(* IEC 61131-3 sources: daoli-st-library/DL_Process (part 24) *)

(* ---- FB_DL_CartonErectSeq.st ---- *)
(*==============================================================================
 * 组件名称 (Component)  : FB_DL_CartonErectSeq
 * 所属子库 (Sublibrary) : DL_Process
 * 当前版本 (Version)    : 1.0.0
 * 兼容性 (Platform)     : CODESYS 3.5 / TwinCAT 3 / 汇川 InoProShop / Machine Expert
 *                         仅依赖纯 IEC 61131-3 标准元素，零厂商方言
 * 功能描述 (Function)   : 开箱机顺控四相：吸箱 → 成型 → 折底 → 输送，含卡箱检测，
 *                         单相超时（tStepMax 默认 5 s）监视；反馈缺失一律进 ERR
 *                         并锁存卡箱（不跳相）；PICK 相真空超时先释放真空再报错；
 *                         CASE 含 ELSE 安全态（全输出 FALSE）；复位退 IDLE。
 * 溯源 (Origin)         : 道莅 clean-room 防御性实现
 * 本文件内含 (Contains) : TYPE E_DL_ErectPhase / TYPE E_DL_ErectErr /
 *                         FUNCTION_BLOCK FB_DL_CartonErectSeq
 * 依赖 (Depends)        : 无 DL_ 内部依赖；Standard.library TON/R_TRIG 实例
 * 红线自检 (Redline)    : 无外部全局变量、无硬件地址直引 ｜ 全变量中英双语同行注释
 *                         相超时用状态判定（TON.Q + 相枚举），非单拍标志 ｜
 *                         枚举成员全部显式赋值 ｜ TON/R_TRIG 每周期无条件调用 ｜
 *                         CASE 含 ELSE 兜底至安全态 ｜ 无占位词 ｜ 超时引脚带单位
 * 错误码表 (Codes)      : 16#0005_041C IDLE（或 DONE 等待下一循环，共用反证句）
 *                         16#0005_041D PICK（吸箱相）
 *                         16#0005_041E FORM（成型相）
 *                         16#0005_041F FLAP（折底相，EJECT 输送段共用反证句）
 *                         16#0005_0420 ERR（含相超时定位，定位另由 eJamPhase 输出）
 * 修订历史 (Revision)   : 2026-11-17  v1.0.0  首版入库 · R27 · 阶段三批 4
 * 验收向量 (Acceptance) : bStart → PICK（真空指令置位）→ bVacuumOk → FORM → bBoxFormed
 *                         → FLAP → bFlapClosed → EJECT → DONE；PICK 相 tStepMax 内
 *                         无 bVacuumOk → ERR + bJam + 真空撤 + eJamPhase=PICK
 *============================================================================*)

(*-----------------------------------------------------------------------------
 * 枚举: E_DL_ErectPhase（归属 DL_Process，开箱顺控相）
 *----------------------------------------------------------------------------*)
TYPE E_DL_ErectPhase :
(
    ePhaseIdle  := 0,    // 空闲待启动 / Idle, waiting for a start
    ePhasePick  := 10,   // 吸箱相（真空建立）/ Pick phase, vacuum build-up
    ePhaseForm  := 20,   // 成型相 / Forming phase
    ePhaseFlap  := 30,   // 折底相 / Flap-closing phase
    ePhaseEject := 40,   // 输送相（定时完成）/ Eject phase, timed
    ePhaseDone  := 50,   // 循环完成（等待下一循环）/ Cycle done, waiting for the next
    ePhaseErr   := 99    // 故障相（卡箱锁存）/ Error phase, jam latched
);
END_TYPE

(*-----------------------------------------------------------------------------
 * 枚举: E_DL_ErectErr（归属 DL_Process，与 FB_DL_CartonErectSeq 同文件）
 *----------------------------------------------------------------------------*)
TYPE E_DL_ErectErr :
(
    eIdle   := 16#0005_041C,   // IDLE（含 DONE 等待态）/ Idle or done-waiting
    ePick   := 16#0005_041D,   // PICK 相（吸箱）/ Pick phase
    eForm   := 16#0005_041E,   // FORM 相（成型）/ Form phase
    eFlap   := 16#0005_041F,   // FLAP 相（折底，含 EJECT 输送段）/ Flap phase, includes eject
    eErr    := 16#0005_0420    // ERR 相（含相超时定位）/ Error phase with timeout localisation
);
END_TYPE

(*==============================================================================
 * 功能块: FB_DL_CartonErectSeq
 * 调用约定: 每个扫描周期无条件调用一次。
 *============================================================================*)
FUNCTION_BLOCK FB_DL_CartonErectSeq
VAR_INPUT
    bVacuumOk    : BOOL;               // 真空建立反馈 / Vacuum established feedback
    bBoxFormed   : BOOL;               // 成型到位反馈 / Box formed feedback
    bFlapClosed  : BOOL;               // 折底到位反馈 / Flap closed feedback
    tStepMax     : TIME := T#5S;       // 单相超时 [秒]，默认 5 / Per-phase timeout [s]
    bStart       : BOOL;               // 启动（上升沿）/ Start, rising edge
    bReset       : BOOL;               // 复位（上升沿，退 IDLE 并清卡箱）/ Reset, rising edge
END_VAR
VAR_OUTPUT
    ePhase       : E_DL_ErectPhase;    // 顺控当前相 / Current sequence phase
    bDone        : BOOL;               // 循环完成（单拍脉冲）/ Cycle done, single-scan pulse
    bJam         : BOOL;               // 卡箱锁存（需复位）/ Jam latched until reset
    eJamPhase    : E_DL_ErectPhase;    // 超时定位相（卡箱时有效）/ Phase where the jam occurred
    bVacuumCmd   : BOOL;               // 真空指令 / Vacuum command
    bConveyorCmd : BOOL;               // 输送指令 / Conveyor command
    eErr         : E_DL_ErectErr;      // 错误码 / Error code
END_VAR
VAR
    fbStartTrig  : R_TRIG;             // 启动沿实例（无条件调用）/ Start edge instance
    fbResetTrig  : R_TRIG;             // 复位沿实例（无条件调用）/ Reset edge instance
    tonStep      : TON;                // 单相超时定时器（无条件调用）/ Per-phase timeout timer
    bPhaseRun    : BOOL;               // 相内计时使能（PICK~EJECT）/ Phase timing enable
END_VAR

(*------------------------------------------------------------------------------
 * 段 1｜沿检测与 TON 每周期无条件调用（仅 IN 条件化）：相超时用状态判定
 *----------------------------------------------------------------------------*)
fbStartTrig(CLK := bStart);                           // 启动沿检测无条件刷新 / start edge refreshed unconditionally
fbResetTrig(CLK := bReset);                           // 复位沿检测无条件刷新 / reset edge refreshed unconditionally
bPhaseRun := (ePhase = E_DL_ErectPhase.ePhasePick) OR (ePhase = E_DL_ErectPhase.ePhaseForm)
          OR (ePhase = E_DL_ErectPhase.ePhaseFlap) OR (ePhase = E_DL_ErectPhase.ePhaseEject);   // 动作相判据 / timed-phase predicate
tonStep(IN := bPhaseRun, PT := tStepMax);             // 单相超时计时（无条件刷新）/ per-phase timing

(*------------------------------------------------------------------------------
 * 段 2｜复位沿：回 IDLE 并清卡箱锁存
 *----------------------------------------------------------------------------*)
IF fbResetTrig.Q THEN
    ePhase := E_DL_ErectPhase.ePhaseIdle;             // 回空闲 / back to idle
    bJam := FALSE;                                    // 卡箱解锁 / jam released
    bDone := FALSE;                                   // 完成撤 / done dropped
    bVacuumCmd := FALSE;                              // 真空撤 / vacuum dropped
    bConveyorCmd := FALSE;                            // 输送撤 / conveyor dropped
    eJamPhase := E_DL_ErectPhase.ePhaseIdle;          // 定位相清 / jam phase cleared
END_IF

(*------------------------------------------------------------------------------
 * 段 3｜启动沿：仅在 IDLE/DONE 允许启动（卡箱态必须复位）
 *----------------------------------------------------------------------------*)
IF fbStartTrig.Q THEN
    IF (ePhase = E_DL_ErectPhase.ePhaseIdle) OR (ePhase = E_DL_ErectPhase.ePhaseDone) THEN
        ePhase := E_DL_ErectPhase.ePhasePick;         // 进吸箱相 / enter pick phase
        bDone := FALSE;                               // 完成撤 / done dropped
    END_IF
END_IF

(*------------------------------------------------------------------------------
 * 段 4｜顺控状态机：CASE 含 ELSE 兜底（ELSE → 安全态全输出 FALSE）
 *----------------------------------------------------------------------------*)
bDone := FALSE;                                       // 完成脉冲逐拍先清 / done pulse cleared first
CASE ePhase OF

    E_DL_ErectPhase.ePhaseIdle:
        bVacuumCmd := FALSE;                          // 空闲：真空撤 / vacuum dropped
        bConveyorCmd := FALSE;                        // 空闲：输送撤 / conveyor dropped
        eErr := E_DL_ErectErr.eIdle;                  // 码 041C / code idle

    E_DL_ErectPhase.ePhasePick:
        bVacuumCmd := TRUE;                           // 吸箱：真空指令置位 / vacuum command set
        bConveyorCmd := FALSE;                        // 吸箱：输送撤 / conveyor dropped
        eErr := E_DL_ErectErr.ePick;                  // 码 041D / code pick
        IF bVacuumOk THEN
            ePhase := E_DL_ErectPhase.ePhaseForm;     // 真空建立：进成型相 / vacuum ok: enter form
        ELSIF tonStep.Q THEN
            bVacuumCmd := FALSE;                      // 真空超时：先释放真空再报错 / vacuum timeout: release vacuum first
            ePhase := E_DL_ErectPhase.ePhaseErr;      // 进故障相 / enter error phase
            bJam := TRUE;                             // 卡箱锁存 / jam latched
            eJamPhase := E_DL_ErectPhase.ePhasePick;  // 定位相 = PICK / jam phase recorded
            eErr := E_DL_ErectErr.eErr;               // 码 0420 / code error
        END_IF

    E_DL_ErectPhase.ePhaseForm:
        bVacuumCmd := TRUE;                           // 成型：真空保持 / vacuum held
        bConveyorCmd := FALSE;                        // 成型：输送撤 / conveyor dropped
        eErr := E_DL_ErectErr.eForm;                  // 码 041E / code form
        IF bBoxFormed THEN
            ePhase := E_DL_ErectPhase.ePhaseFlap;     // 成型到位：进折底相 / formed: enter flap
        ELSIF tonStep.Q THEN
            bVacuumCmd := FALSE;                      // 超时：撤真空（安全侧）/ timeout: drop vacuum
            ePhase := E_DL_ErectPhase.ePhaseErr;      // 进故障相 / enter error
            bJam := TRUE;                             // 卡箱锁存 / jam latched
            eJamPhase := E_DL_ErectPhase.ePhaseForm;  // 定位相 = FORM / jam phase recorded
            eErr := E_DL_ErectErr.eErr;               // 码 0420 / code error
        END_IF

    E_DL_ErectPhase.ePhaseFlap:
        bVacuumCmd := TRUE;                           // 折底：真空保持 / vacuum held
        bConveyorCmd := FALSE;                        // 折底：输送撤 / conveyor dropped
        eErr := E_DL_ErectErr.eFlap;                  // 码 041F / code flap
        IF bFlapClosed THEN
            ePhase := E_DL_ErectPhase.ePhaseEject;    // 折底到位：进输送相 / flap closed: enter eject
        ELSIF tonStep.Q THEN
            bVacuumCmd := FALSE;                      // 超时：撤真空（安全侧）/ timeout: drop vacuum
            ePhase := E_DL_ErectPhase.ePhaseErr;      // 进故障相 / enter error
            bJam := TRUE;                             // 卡箱锁存 / jam latched
            eJamPhase := E_DL_ErectPhase.ePhaseFlap;  // 定位相 = FLAP / jam phase recorded
            eErr := E_DL_ErectErr.eErr;               // 码 0420 / code error
        END_IF

    E_DL_ErectPhase.ePhaseEject:
        bVacuumCmd := FALSE;                          // 输送：真空撤（放箱）/ eject: vacuum dropped
        bConveyorCmd := TRUE;                         // 输送：输送指令置位 / conveyor command set
        eErr := E_DL_ErectErr.eFlap;                  // 码 041F（输送段与折底段共用，反证句见文件头）/ code flap, shared band
        IF tonStep.Q THEN
            bConveyorCmd := FALSE;                    // 输送定时到：撤输送 / timed eject: drop conveyor
            bDone := TRUE;                            // 完成单拍脉冲 / single-scan done pulse
            ePhase := E_DL_ErectPhase.ePhaseDone;     // 进完成相 / enter done
        END_IF

    E_DL_ErectPhase.ePhaseDone:
        bVacuumCmd := FALSE;                          // 完成：真空撤 / vacuum dropped
        bConveyorCmd := FALSE;                        // 完成：输送撤 / conveyor dropped
        eErr := E_DL_ErectErr.eIdle;                  // 码 041C（DONE 等待态与 IDLE 输出组合相同，共用反证句）/ code idle, shared band

    E_DL_ErectPhase.ePhaseErr:
        bVacuumCmd := FALSE;                          // 故障相：真空撤 / vacuum dropped
        bConveyorCmd := FALSE;                        // 故障相：输送撤 / conveyor dropped
        bJam := TRUE;                                 // 卡箱保持锁存 / jam held latched
        eErr := E_DL_ErectErr.eErr;                   // 码 0420 / code error

    ELSE
        ePhase := E_DL_ErectPhase.ePhaseErr;          // 非法相兜底 / illegal-phase fallback
        bVacuumCmd := FALSE;                          // 安全态：真空撤 / vacuum dropped, safe side
        bConveyorCmd := FALSE;                        // 安全态：输送撤 / conveyor dropped, safe side
        bJam := TRUE;                                 // 卡箱锁存（非法相按卡箱处置）/ jam latched
        eJamPhase := E_DL_ErectPhase.ePhaseErr;       // 定位相 = ERR / jam phase recorded
        eErr := E_DL_ErectErr.eErr;                   // 码 0420 / code error

END_CASE
END_FUNCTION_BLOCK

(* ---- FB_DL_CartonScannerSort.st ---- *)
(*
  Component : FB_DL_CartonScannerSort
  Category  : DL_Process
  Type      : FB
  Version   : 1.0.0
  CodeSeg   : 16#06_0_3C
  Summary   : 纸箱扫码分道：读码判定 + 分道放行调度（与输送段 Zone 握手防追尾），读码失败走旁路 NG 道。
              Carton scanner sort: read verdict plus lane dispatch with zone handshake, read fail bypasses to the NG lane.
  溯源声明  : 道莅自研 clean-room
  边界安全  : 与 FB_DL_ConveyorZone 段间握手经 VAR_IN_OUT（ioZoneFree / ioDispatchAck），不写对方内部状态；
              步进超时 tAckMs 提为输入引脚，超时回安全步（NG 旁路，不堵线）；条码号负值域拦截；
              分道放行单拍脉冲防重复放行；CASE 必带 ELSE 安全步；TON 每拍无条件刷新。
  复用      : 与 FB_DL_ConveyorZone 握手（VAR_IN_OUT 引脚级，无实例依赖）；复用 FB_DL_StepSequencer 步进语义（clean-room 自含实现）
*)

FUNCTION_BLOCK FB_DL_CartonScannerSort
VAR_INPUT
    bRun      : BOOL;                   (* 调度使能 · Enable *)
    bScanTrig : BOOL;                   (* 扫码触发 [事件]，到位传感器 · Scan trigger pulse *)
    bReadOk   : BOOL;                   (* 读码成功反馈 [开关] · Read success feedback *)
    nCode     : DINT;                   (* 条码号 [号]，负值拦截 · Barcode number *)
    nLaneCnt  : INT := 3;               (* 合格分道数 [道]，域 1 到 3 · OK lane count *)
    tAckMs    : TIME  := T#2000MS;      (* 放行应答超时 [ms] · Dispatch ack timeout *)
    fEps      : LREAL := 1.0E-6;        (* 浮点判零容差 [实数域] · Floating zero tolerance *)
END_VAR
VAR_IN_OUT
    ioZoneFree    : BOOL;               (* 上游 Zone 空闲握手 [引脚] · Zone free handshake *)
    ioDispatchAck : BOOL;               (* 分道执行应答 [引脚]，由 Zone 件置位 · Dispatch ack from zone *)
END_VAR
VAR_OUTPUT
    eStep    : (eStpWait := 0, eStpDispatch := 1, eStpAck := 2);     (* 步枚举输出 / Step output enum *)
    nLaneSel : INT;                     (* 选中道号 [道]，1 到 nLaneCnt，0 为 NG 旁路 · Selected lane *)
    bDispatch: BOOL;                    (* 分道放行脉冲 [脉冲] · Dispatch pulse *)
    nOkCount : UDINT;                   (* 合格道累计 [件]，防回卷 · OK count *)
    nNgCount : UDINT;                   (* NG 旁路累计 [件]，防回卷 · NG count *)
    bError   : BOOL;                    (* 故障标志，与故障码配对 · Fault flag paired with codes *)
    uErrorId : UDINT;                   (* 事件码 16#0000_003C，0 无事件 · Event code *)
END_VAR
VAR
    _eState : (eStWait := 0, eStDispatch := 1, eStAck := 2);    (* 内部步进状态 / Internal step state *)
    uCode   : WORD;     (* 码位暂存，每拍重算 [码] · Code staging *)
    tonAck  : TON;      (* 应答超时计时 [ms]，每拍无条件刷新 · Ack timeout timer *)
    bTrigPrv: BOOL;     (* 上拍触发快照，上升沿判据 · Previous trigger snapshot *)
    bTrig   : BOOL;     (* 扫码上升沿 [脉冲] · Scan rising edge *)
    nCycles : UDINT;    (* 分道累计 [件]，防回卷 · Dispatch count *)
END_VAR
VAR CONSTANT
    DL_CSS_WRAP : UDINT := 4294967290;  (* 计数防回卷余量 [件] · Counter wrap guard *)
END_VAR

(* === 段 0 · 实例刷新（每拍无条件，红线 7）=== *)
tonAck(IN := (_eState = eStAck), PT := tAckMs);     (* 应答超时计时 / Ack timeout timing *)
bTrig := bScanTrig AND (NOT bTrigPrv);              (* 扫码上升沿 / Scan rising edge *)
bTrigPrv := bScanTrig;                              (* 快照更新 / Snapshot *)

(* === 段 1 · 输入校验与量程闸 === *)
uCode := 16#0000;                       // 每拍清码（可达清零基线）/ Clear codes each scan
IF (nLaneCnt < 1) OR (nLaneCnt > 3) OR (tAckMs <= T#0MS) THEN
    uCode := 16#003C;                   // 故障级：整定域外，调度冻结 / Fault: tuning domain invalid
END_IF

(* === 段 2 · 主逻辑：步进状态机（步进 CASE 必带 ELSE 安全步）=== *)
CASE _eState OF
    eStWait:                            (* 等待步：触发且 Zone 空闲才进入分派 / Wait for trigger and zone *)
        nLaneSel := 0;                  (* 道号清零待选 / Clear lane selection *)
        bDispatch := FALSE;             (* 放行脉冲收口 / Dispatch pulse off *)
        IF bRun AND (uCode = 16#0000) AND bTrig AND ioZoneFree THEN
            _eState := eStDispatch;     (* 拍 N 条件满足，拍 N+1 分派 / To dispatch next scan *)
        END_IF
    eStDispatch:                        (* 分派步：读码判定选道，失败走 NG 旁路不堵线 / Select lane, fail bypasses *)
        IF bReadOk AND (nCode >= 0) THEN
            nLaneSel := (UDINT_TO_DINT(INT_TO_UDINT(1)) + (nCode MOD UDINT_TO_DINT(INT_TO_UDINT(nLaneCnt))));
                                        (* 均衡选道：1 + 条码 mod 道数 / Balanced lane pick *)
            IF nOkCount < DL_CSS_WRAP THEN
                nOkCount := nOkCount + 1;   (* 合格计数 / Count OK *)
            END_IF
        ELSE
            nLaneSel := 0;              (* 读码失败：NG 旁路道 / Read fail: NG bypass lane *)
            IF nNgCount < DL_CSS_WRAP THEN
                nNgCount := nNgCount + 1;   (* NG 计数 / Count NG *)
            END_IF
        END_IF
        bDispatch := TRUE;              (* 放行脉冲发出 / Issue the dispatch pulse *)
        _eState := eStAck;              (* 拍 N 分派，拍 N+1 等应答 / To ack next scan *)
    eStAck:                             (* 应答步：应答回等待，超时安全步 / Await ack, timeout to safe step *)
        bDispatch := FALSE;             (* 脉冲单拍收口 / One-scan pulse off *)
        IF ioDispatchAck THEN
            _eState := eStWait;         (* 应答确认回等待 / Acked back to wait *)
        ELSIF tonAck.Q THEN
            _eState := eStWait;         (* 超时回安全等待步（NG 旁路语义，不堵线）/ Timeout to safe step *)
            uCode := 16#003C;           (* 故障级：应答超时 / Fault: ack timeout *)
        END_IF
ELSE
    _eState := eStWait;                 (* ELSE 兜底回安全等待步 / ELSE fallback to safe step *)
    bDispatch := FALSE;
    nLaneSel := 0;
END_CASE

(* === 段 3 · 输出映射与故障码（CASE 内未触碰输出枚举）=== *)
eStep := eStpWait;                      (* 步映射默认 / Default mapping *)
IF _eState = eStDispatch THEN
    eStep := eStpDispatch;              (* 分派步映射 / Map dispatch *)
ELSIF _eState = eStAck THEN
    eStep := eStpAck;                   (* 应答步映射 / Map ack *)
END_IF
IF nOkCount + nNgCount > DL_CSS_WRAP THEN
    nCycles := nOkCount + nNgCount;     (* 分道累计与两计数口径对齐 / Align the dispatch ledger *)
END_IF
bError := (uCode <> 16#0000);           (* 故障标志配对 / Fault flag paired *)
uErrorId := WORD_TO_UDINT(uCode);       (* 码位单点写入（16#0000_003C 形态）/ Single write point *)
END_FUNCTION_BLOCK

(* ---- FB_DL_CasePackerPattern.st ---- *)
//==============================================================================
// 功能块：FB_DL_CasePackerPattern ｜ 中文名称：装箱排列模式生成
// 所属子库：DL_Process ｜ 版本：v1.0.0 ｜ 兼容：CODESYS V3.5+ / TwinCAT 3 / 汇川 InoProShop
// 功能描述：装箱机的排列模式生成件：按箱型规格（列数 / 行数 / 层数 / 节距 / 交错方式）
//           把「盒号」解码成「目标位姿 X/Y/Z + 旋转标志」的抓取序列，支持行交错（奇数行
//           半节距平移）与整层 90 度旋转（层号循环 0/90/180/270，旋转层 X/Y 轴互换）。
//           本件只生成序列与握手位，不执行任何动作、不驱动机器人、不做轨迹规划（位姿
//           给到上层定位层）。序号推进用 bStepDone 握手位的上升沿：上层置位表示本步已
//           执行完毕，本件取沿推进并自清（单拍标志自清，防同一格位重复取件）。
// 开源溯源 (Origin)：道莅原创实现（参考 公开工程惯例 分类与参数域）
// 单位表：节距/层距/坐标[mm] / 旋转角[度] / 行列层[个] / 槽位与盒数[件]
// 错误码表：16#0005_0404 信息级（装箱容量大于本箱数量，末层留空位，不置 bError）/
//           16#0005_0405 信息级（交错/层旋转配置与单层配置冲突被规格钳位为无交错，
//           不置 bError）/ 16#0005_0348 故障级（排列容量小于本箱数量，或行列层域外
//           1~20，或数量域非法，置 bError）/ 16#0005_0349 故障级（节距/层距非正或任一
//           浮点输入非有限，置 bError——尺寸非法与非有限共用本槽，反证句：二者在现有
//           输出组合下不可观测出差异，均为 bValid 撤 + 序列回序号 1）/ 16#0005_034A
//           故障级兜底（状态机落 ELSE 非法状态，置 bError）。码位 16#0005 段。
// 状态机：E_DL_CasePackState（eIdle=0 待机 / eRunning=10 序列输出中 / eDone=20 末位已
//           输出 / eFault=99 故障兜底），CASE 含 ELSE 兜底，ELSE 置 034A 且序列回 1、
//           许可撤。
// 边界行为：① 容量 nCols x nRows x nLayers 与 nBoxCount 校验：nBoxCount > 容量 → 故障
//           0348（绝不硬塞）；nBoxCount < 容量 → 合法（末层留空位）+ 信息 0404 +
//           nEmptySlots 出口；② 行列层域外（≤ 0 或 > 20）→ 故障 0348；③ 节距 ≤ 0 或
//           非有限 → 故障 0349（防负坐标倒排、防非有限坐标外泄）；④ 序列越界防护：
//           nSeqIndex 达 nBoxCount 即 bLast 且不再推进；⑤ nLayers = 1 且 eLayerRotate
//           → 钳为 eNone + 信息 0405；⑥ 失能 → 序列复位到序号 1 + bValid := FALSE
//           （R72）；⑦ 坐标解算只做乘加与整除，除子为已判正的行列数（先判后除）。
// 修订历史：v1.0.0 2026-11-17 首版（R25 派单 · §4.14）
//==============================================================================
(*------------------------------------------------------------------------------
 * 枚举: E_DL_PackInterlock（归属 DL_Process，与 FB_DL_CasePackerPattern 同文件）
 *       装箱交错方式；数值步长留空位，便于后续插值不破坏已有工程
 *----------------------------------------------------------------------------*)
TYPE E_DL_PackInterlock :
(
    eNone        := 0,   // 无交错：行列正交直排 / No interlock, orthogonal grid
    eRowShift    := 10,  // 行交错：奇数行沿列方向平移半个节距 / Row interlock, odd rows shifted half a pitch
    eLayerRotate := 20   // 层旋转：逐层循环旋转 0/90/180/270 度 / Layer rotation cycling 0/90/180/270 degrees
);
END_TYPE

(*------------------------------------------------------------------------------
 * 枚举: E_DL_CasePackState（归属 DL_Process，与 FB_DL_CasePackerPattern 同文件）
 *----------------------------------------------------------------------------*)
TYPE E_DL_CasePackState :
(
    eIdle    := 0,   // 待机：序列复位到序号 1，许可撤 / Idle, sequence reset to index 1, permission dropped
    eRunning := 10,  // 输出中：逐盒给出目标位姿 / Running, target pose emitted per case
    eDone    := 20,  // 末位已输出：bLast 置位，等待复位 / Last slot emitted, waiting for reset
    eFault   := 99   // 故障兜底：规格非法/非有限/非法状态 / Fault fallback
);
END_TYPE

(*==============================================================================
 * 功能块: FB_DL_CasePackerPattern
 * 调用约定: 每个扫描周期无条件调用一次；上层在完成一次抓取后把 bStepDone 置 TRUE。
 *============================================================================*)
FUNCTION_BLOCK FB_DL_CasePackerPattern
VAR_INPUT
    nCols          : INT;                          // 列数 [个]，合法域 1~20 / Column count [pcs], domain 1..20
    nRows          : INT;                          // 行数 [个]，合法域 1~20 / Row count [pcs], domain 1..20
    nLayers        : INT;                          // 层数 [个]，合法域 1~20 / Layer count [pcs], domain 1..20
    fPitchXMm      : LREAL;                        // 列方向节距 [mm]，须 > 0 / Column pitch [mm], must be > 0
    fPitchYMm      : LREAL;                        // 行方向节距 [mm]，须 > 0 / Row pitch [mm], must be > 0
    fLayerGapMm    : LREAL;                        // 层间高度差 [mm]，须 > 0 / Layer height gap [mm], must be > 0
    eInterlock     : E_DL_PackInterlock;           // 交错方式（无 / 行交错 / 层旋转）/ Interlock mode
    nBoxCount      : INT;                          // 本箱数量 [件]，合法域 1~容量 / Cases in this carton [pcs], domain 1..capacity
    bEnable        : BOOL;                         // 总使能 / Master enable
    bReset         : BOOL;                         // 复位，上升沿把序列复位到序号 1 / Reset, rising edge rewinds the sequence to index 1
END_VAR
VAR_OUTPUT
    nSeqIndex      : INT;                          // 当前序号 [个]，从 1 起 / Current sequence index, 1-based
    fTargetXMm     : LREAL;                        // 目标位 X [mm] / Target X [mm]
    fTargetYMm     : LREAL;                        // 目标位 Y [mm] / Target Y [mm]
    fTargetZMm     : LREAL;                        // 目标位 Z [mm]，按层高累计 / Target Z [mm], accumulated per layer
    fTargetRotDeg  : LREAL;                        // 目标旋转角 [度]，取 0 / 90 / 180 / 270 / Target rotation [deg], 0/90/180/270
    bStepDone      : BOOL;                         // 本步完成握手位（上层置 TRUE，本件取沿后自清）/ Step handshake, caller sets TRUE, the block clears it after consuming
    bLast          : BOOL;                         // 末位标志（本箱最后一个非空槽位）/ Last slot of this carton
    nSlotCount     : INT;                          // 总槽位数 [件] = 列 x 行 x 层 / Total slots [pcs]
    nEmptySlots    : INT;                          // 空槽位数 [件] = 总槽位 − 本箱数量 / Empty slots [pcs]
    eErr           : UDINT;                        // 错误码，0 = 无错，码位 16#0005_0404 起信息级、16#0005_0348 起故障级（分带见错误码表） / Error code, 0 = no error, band info/fault per the code table
    bError         : BOOL;                         // 故障级标志，仅故障级错误置位 / Fault-class flag, set only on fault-level codes
    bValid         : BOOL;                        // 位姿输出可用标志，失能/故障闸显式 FALSE / Pose usable flag, explicit FALSE on disable/fault gates
    eState         : E_DL_CasePackState;           // 主状态机当前状态 / Current state of the main state machine
END_VAR
VAR
    fbReset        : R_TRIG;                       // 复位上升沿检测实例 / Reset rising edge detector
    fbStep         : R_TRIG;                       // 步完成握手上升沿检测实例 / Step handshake rising edge detector
    eInterlockEff  : E_DL_PackInterlock;           // 生效交错方式（钳位后）/ Effective interlock mode after clamping
    nCapacity      : INT;                          // 总容量 [件] = 列 x 行 x 层 / Total capacity [pcs]
    nIdx0          : INT;                          // 零基序号 [—] / Zero-based sequence index
    nPerLayer      : INT;                          // 每层盒数 [件] = 列 x 行 / Cases per layer [pcs]
    nLayer         : INT;                          // 层号（1 基）[层] / Layer number, 1-based
    nRemain        : INT;                          // 层内余量序号 [—] / In-layer remainder index
    nRow           : INT;                          // 行号（1 基）[行] / Row number, 1-based
    nCol           : INT;                          // 列号（1 基）[列] / Column number, 1-based
    nRotQuarter    : INT;                          // 旋转四分之一圈数 [—] / Rotation quarter count
    fShiftXMm      : LREAL;                        // 行交错平移量 [mm] / Row interlock shift [mm]
    bClampInterlock : BOOL;                        // 交错配置被钳位标志 / Interlock clamped flag
    bSpaceWarn     : BOOL;                         // 末层留空位提示标志 / Empty-slot hint flag
    bFirstScan     : BOOL := TRUE;                 // 上电首拍标志 / First-scan flag
END_VAR
VAR CONSTANT
    DL_CPP_CODE_INFO_1 : UDINT := 16#0005_0404;    // 信息级槽 1（容量大于数量，末层留空位） / info slot 1
    DL_CPP_CODE_INFO_2 : UDINT := 16#0005_0405;    // 信息级槽 2（交错/层旋转配置被钳位） / info slot 2
    DL_CPP_CODE_FLT_1  : UDINT := 16#0005_0348;    // 故障级槽 1（容量不足/行列层域非法） / fault slot 1
    DL_CPP_CODE_FLT_2  : UDINT := 16#0005_0349;    // 故障级槽 2（尺寸非法/输入非有限） / fault slot 2
    DL_CPP_CODE_FLT_3  : UDINT := 16#0005_034A;    // 故障级槽 3（非法状态兜底） / fault slot 3, illegal-state fallback
    DL_CPP_DIM_MIN     : INT := 1;                 // 行列层下限 [个] / Dimension floor [pcs]
    DL_CPP_DIM_MAX     : INT := 20;                // 行列层上限 [个] / Dimension ceiling [pcs]
    DL_CPP_ZERO        : LREAL := 0.0;             // 零值常量，避免裸字面量 [—] / Zero constant, avoids a bare literal
    DL_CPP_TOL         : LREAL := 1.0E-6;          // 浮点比较容差 [—] / Float comparison tolerance
    DL_CPP_INF         : LREAL := 1.7976931348623157E308; // LREAL 幅值上限，Inf 判据 / LREAL magnitude ceiling
    DL_CPP_HALF        : LREAL := 0.5;             // 半节距系数 [—] / Half-pitch factor
    DL_CPP_QUARTER_DEG : LREAL := 90.0;            // 每层旋转步长 [度] / Rotation step per layer [deg]
    DL_CPP_QUARTERS    : INT := 4;                 // 旋转循环周期 [层] / Rotation cycle length [layers]
    DL_CPP_IDX_FIRST   : INT := 1;                 // 序号起点 [个] / First sequence index
END_VAR

(*------------------------------------------------------------------------------
 * 段 1｜无条件刷新区（红线 5）：复位沿与步完成握手沿在任意分支之外周期调用
 *----------------------------------------------------------------------------*)
fbReset(CLK := bReset);                            // 复位沿检测无条件刷新 / reset edge refreshed unconditionally
fbStep(CLK := bStepDone);                          // 步完成沿检测无条件刷新（先取沿后自清）/ step edge refreshed before the output is cleared

(*------------------------------------------------------------------------------
 * 段 2｜复位沿处理（改写置于沿后，防吞沿 R39）
 *----------------------------------------------------------------------------*)
IF fbReset.Q THEN
    eState := E_DL_CasePackState.eIdle;
    eErr   := 16#0000_0000;                        // 复位清码 / reset clears the code
    bError := FALSE;                               // 复位清故障 / reset clears the fault
    nSeqIndex := DL_CPP_IDX_FIRST;                 // 序列复位到序号 1 / sequence rewound to index 1
    bStepDone := FALSE;                            // 握手位清 / handshake cleared
    bFirstScan := TRUE;                            // 重新首拍化 / re-initialize first scan
END_IF

(*------------------------------------------------------------------------------
 * 段 3｜非有限输入闸：尺寸类浮点非有限 → 0349（与尺寸非法共用本槽，见头注释反证句）
 *----------------------------------------------------------------------------*)
IF (fPitchXMm <> fPitchXMm) OR (ABS(fPitchXMm) >= DL_CPP_INF)
   OR (fPitchYMm <> fPitchYMm) OR (ABS(fPitchYMm) >= DL_CPP_INF)
   OR (fLayerGapMm <> fLayerGapMm) OR (ABS(fLayerGapMm) >= DL_CPP_INF) THEN
    eState := E_DL_CasePackState.eFault;           // 进故障相 / enter fault state
    eErr   := DL_CPP_CODE_FLT_2;                   // 故障级：输入非有限 / fault: non-finite input
    bError := TRUE;                                // 故障级必置 bError（R45 配对）/ fault-class pairs with bError
    bValid := FALSE;                               // 位姿不可用 / poses unusable
    nSeqIndex := DL_CPP_IDX_FIRST;                 // 序列回序号 1 安全侧 / sequence rewound, safe side
    fTargetXMm := DL_CPP_ZERO;                     // 坐标回零安全侧 / coordinates zeroed, safe side
    fTargetYMm := DL_CPP_ZERO;                     // 坐标回零安全侧 / coordinates zeroed, safe side
    fTargetZMm := DL_CPP_ZERO;                     // 坐标回零安全侧 / coordinates zeroed, safe side
    fTargetRotDeg := DL_CPP_ZERO;                  // 旋转角回零安全侧 / rotation zeroed, safe side
    bLast := FALSE;                                // 末位标志撤 / last flag withdrawn
    RETURN;
END_IF

(*------------------------------------------------------------------------------
 * 段 4｜组态合法性闸：行列层域（1~20）+ 节距层距为正（防负坐标倒排、防除零）
 *----------------------------------------------------------------------------*)
IF (nCols < DL_CPP_DIM_MIN) OR (nCols > DL_CPP_DIM_MAX)
   OR (nRows < DL_CPP_DIM_MIN) OR (nRows > DL_CPP_DIM_MAX)
   OR (nLayers < DL_CPP_DIM_MIN) OR (nLayers > DL_CPP_DIM_MAX) THEN
    eState := E_DL_CasePackState.eFault;           // 进故障相 / enter fault state
    eErr   := DL_CPP_CODE_FLT_1;                   // 故障级：行列层域非法 / fault: dimension out of range
    bError := TRUE;                                // 故障级必置 bError（R45 配对）/ fault-class pairs with bError
    bValid := FALSE;                               // 位姿不可用 / poses unusable
    nSeqIndex := DL_CPP_IDX_FIRST;                 // 序列回序号 1 安全侧 / sequence rewound, safe side
    fTargetXMm := DL_CPP_ZERO;                     // 坐标回零安全侧 / coordinates zeroed, safe side
    fTargetYMm := DL_CPP_ZERO;                     // 坐标回零安全侧 / coordinates zeroed, safe side
    fTargetZMm := DL_CPP_ZERO;                     // 坐标回零安全侧 / coordinates zeroed, safe side
    fTargetRotDeg := DL_CPP_ZERO;                  // 旋转角回零安全侧 / rotation zeroed, safe side
    bLast := FALSE;                                // 末位标志撤 / last flag withdrawn
    RETURN;
END_IF
IF (fPitchXMm <= DL_CPP_TOL) OR (fPitchYMm <= DL_CPP_TOL) OR (fLayerGapMm <= DL_CPP_TOL) THEN
    eState := E_DL_CasePackState.eFault;           // 进故障相 / enter fault state
    eErr   := DL_CPP_CODE_FLT_2;                   // 故障级：尺寸非法 / fault: dimension invalid
    bError := TRUE;                                // 故障级必置 bError（R45 配对）/ fault-class pairs with bError
    bValid := FALSE;                               // 位姿不可用 / poses unusable
    nSeqIndex := DL_CPP_IDX_FIRST;                 // 序列回序号 1 安全侧 / sequence rewound, safe side
    fTargetXMm := DL_CPP_ZERO;                     // 坐标回零安全侧 / coordinates zeroed, safe side
    fTargetYMm := DL_CPP_ZERO;                     // 坐标回零安全侧 / coordinates zeroed, safe side
    fTargetZMm := DL_CPP_ZERO;                     // 坐标回零安全侧 / coordinates zeroed, safe side
    fTargetRotDeg := DL_CPP_ZERO;                  // 旋转角回零安全侧 / rotation zeroed, safe side
    bLast := FALSE;                                // 末位标志撤 / last flag withdrawn
    RETURN;
END_IF

(*------------------------------------------------------------------------------
 * 段 5｜容量自算与数量校验：容量不足绝不硬塞（0348），容量富余属合法（0404）
 *----------------------------------------------------------------------------*)
nCapacity := nCols * nRows * nLayers;              // 总容量 [件] / total capacity [pcs]
nPerLayer := nCols * nRows;                        // 每层盒数 [件] / cases per layer [pcs]
nSlotCount := nCapacity;                           // 总槽位出口 / total slot count outlet
IF (nBoxCount < DL_CPP_DIM_MIN) OR (nBoxCount > nCapacity) THEN
    eState := E_DL_CasePackState.eFault;           // 进故障相 / enter fault state
    eErr   := DL_CPP_CODE_FLT_1;                   // 故障级：数量域非法或容量不足 / fault: count out of range or capacity exceeded
    bError := TRUE;                                // 故障级必置 bError（R45 配对）/ fault-class pairs with bError
    bValid := FALSE;                               // 位姿不可用 / poses unusable
    nEmptySlots := nCapacity - nBoxCount;          // 空位数为负则如实透出（诊断用）/ empty slots reported even when negative, for diagnosis
    nSeqIndex := DL_CPP_IDX_FIRST;                 // 序列回序号 1 安全侧 / sequence rewound, safe side
    RETURN;
END_IF
nEmptySlots := nCapacity - nBoxCount;              // 空槽位数 [件] / empty slots [pcs]
bSpaceWarn := (nEmptySlots > 0);                   // 末层留空位提示 / empty-slot hint

(*------------------------------------------------------------------------------
 * 段 6｜交错方式钳位：单层配置下的层旋转无意义，钳为无交错（0405）；
 *       枚举越界值同样钳为无交错并提示，不新增码位
 *----------------------------------------------------------------------------*)
eInterlockEff := eInterlock;                       // 先取引脚值 / take the pin value first
bClampInterlock := FALSE;                          // 钳位标志逐拍重判 / clamp flag re-judged per scan
IF (eInterlockEff <> E_DL_PackInterlock.eNone)
   AND (eInterlockEff <> E_DL_PackInterlock.eRowShift)
   AND (eInterlockEff <> E_DL_PackInterlock.eLayerRotate) THEN
    eInterlockEff := E_DL_PackInterlock.eNone;     // 枚举越界：钳为无交错 / out-of-range enumeration clamped to none
    bClampInterlock := TRUE;                       // 钳位提示 / clamp hint
END_IF
IF (eInterlockEff = E_DL_PackInterlock.eLayerRotate) AND (nLayers <= 1) THEN
    eInterlockEff := E_DL_PackInterlock.eNone;     // 单层无层旋转可言 / layer rotation is meaningless with a single layer
    bClampInterlock := TRUE;                       // 钳位提示 / clamp hint
END_IF

(*------------------------------------------------------------------------------
 * 段 7｜握手推进：bStepDone 上升沿推进序号；末位不再推进（序列越界防护）
 *----------------------------------------------------------------------------*)
IF fbStep.Q THEN
    bStepDone := FALSE;                            // 握手位自清（单拍标志自清，红线 5）/ handshake self-cleared
    IF nSeqIndex < nBoxCount THEN
        nSeqIndex := nSeqIndex + 1;                // 推进到下一盒号 / advance to the next case
    END_IF
END_IF
IF nSeqIndex < DL_CPP_IDX_FIRST THEN
    nSeqIndex := DL_CPP_IDX_FIRST;                 // 序号下限防护 / index floor guard
END_IF
IF nSeqIndex > nBoxCount THEN
    nSeqIndex := nBoxCount;                        // 序号上限防护 / index ceiling guard
END_IF
bLast := (nSeqIndex >= nBoxCount);                 // 末位标志（本箱最后一个非空槽位）/ last slot of this carton

(*------------------------------------------------------------------------------
 * 段 8｜盒号解码：零基序号 → 层 / 行 / 列（除子 nPerLayer 与 nCols 已由段 4 保证为正）
 *----------------------------------------------------------------------------*)
nIdx0 := nSeqIndex - DL_CPP_IDX_FIRST;             // 零基序号 / zero-based index
nLayer := (nIdx0 / nPerLayer) + 1;                 // 层号（1 基）[层] / layer number, 1-based
nRemain := nIdx0 - ((nLayer - 1) * nPerLayer);     // 层内余量（显式减法，避开 MOD 的负数方言差异）/ in-layer remainder
nRow := (nRemain / nCols) + 1;                     // 行号（1 基）[行] / row number, 1-based
nCol := nRemain - ((nRow - 1) * nCols) + 1;        // 列号（1 基）[列] / column number, 1-based

(*------------------------------------------------------------------------------
 * 段 9｜位姿解算：层旋转 exch 轴序，行交错平移半节距；Z 按层高累计
 *----------------------------------------------------------------------------*)
fShiftXMm := DL_CPP_ZERO;                          // 交错平移量初值 / interlock shift seed
IF eInterlockEff = E_DL_PackInterlock.eRowShift THEN
    IF ((nRow - 1) MOD 2) = 1 THEN
        fShiftXMm := fPitchXMm * DL_CPP_HALF;      // 奇数行平移半节距 [mm] / odd rows shifted half a pitch
    END_IF
END_IF
nRotQuarter := 0;                                  // 旋转四分之一圈数初值 / rotation quarter seed
IF eInterlockEff = E_DL_PackInterlock.eLayerRotate THEN
    nRotQuarter := (nLayer - 1) MOD DL_CPP_QUARTERS;   // 逐层循环 0/1/2/3 个四分之一圈 / per-layer quarter cycle
END_IF
fTargetRotDeg := INT_TO_LREAL(nRotQuarter) * DL_CPP_QUARTER_DEG;   // 目标旋转角 [度] / target rotation [deg]
IF (nRotQuarter = 1) OR (nRotQuarter = 3) THEN
    fTargetXMm := (INT_TO_LREAL(nRow - 1) * fPitchYMm) + fShiftXMm;   // 旋转层：X 走行方向节距 [mm] / rotated layer, X follows the row pitch
    fTargetYMm := INT_TO_LREAL(nCol - 1) * fPitchXMm;                 // 旋转层：Y 走列方向节距 [mm] / rotated layer, Y follows the column pitch
ELSE
    fTargetXMm := (INT_TO_LREAL(nCol - 1) * fPitchXMm) + fShiftXMm;   // 正交层：X 走列方向节距 [mm] / orthogonal layer, X follows the column pitch
    fTargetYMm := INT_TO_LREAL(nRow - 1) * fPitchYMm;                 // 正交层：Y 走行方向节距 [mm] / orthogonal layer, Y follows the row pitch
END_IF
fTargetZMm := INT_TO_LREAL(nLayer - 1) * fLayerGapMm;                 // 层高累计（LREAL 承载）[mm] / layer height accumulation

(*------------------------------------------------------------------------------
 * 段 10｜状态机：CASE 含 ELSE 兜底（非法状态 → 034A + 序列回 1 + 许可撤）
 *----------------------------------------------------------------------------*)
CASE eState OF

    E_DL_CasePackState.eIdle:
        bValid := FALSE;                           // 失能闸显式不可用（R72）/ explicit FALSE on the disable gate
        nSeqIndex := DL_CPP_IDX_FIRST;             // 待机序列固守序号 1 / idle holds index 1
        bLast := (nBoxCount <= DL_CPP_IDX_FIRST);  // 单件箱待机即末位 / a single-case carton is already last
        eErr := 16#0000_0000;                      // 待机无错 / no error in idle
        bError := FALSE;                           // 待机无故障 / no fault in idle
        IF bEnable THEN
            eState := E_DL_CasePackState.eRunning; // 使能进输出相 / enable enters the running state
            bFirstScan := FALSE;                   // 首拍标志清除 / first-scan flag cleared
        END_IF

    E_DL_CasePackState.eRunning:
        bValid := TRUE;                            // 位姿可用 / poses usable
        bError := FALSE;                           // 输出相无故障 / no fault in the running state
        eErr := 16#0000_0000;                      // 输出相先清码 / clear the code first
        IF bClampInterlock THEN
            eErr := DL_CPP_CODE_INFO_2;            // 信息级：交错配置被钳位 / info: interlock clamped
        END_IF
        IF bSpaceWarn THEN
            eErr := DL_CPP_CODE_INFO_1;            // 信息级：末层留空位（与钳位提示并列时以空位为主）/ info: empty slots, the primary hint
        END_IF
        IF NOT bEnable THEN
            eState := E_DL_CasePackState.eIdle;    // 失能回待机（退出条件一）/ disable, first exit
            bValid := FALSE;                       // 失能闸显式不可用 / explicit FALSE on the disable gate
            nSeqIndex := DL_CPP_IDX_FIRST;         // 序列复位到序号 1 / sequence rewound
        ELSIF bLast AND fbStep.Q THEN
            eState := E_DL_CasePackState.eDone;    // 末位已完成转完成相（退出条件二）/ last slot done, second exit
        END_IF

    E_DL_CasePackState.eDone:
        bValid := TRUE;                            // 末位位姿仍可读（现场常需复核）/ the last pose stays readable
        bLast := TRUE;                             // 末位标志保持 / last flag held
        bError := FALSE;                           // 完成相无故障 / no fault in the done state
        eErr := DL_CPP_CODE_INFO_1;                // 信息级：末层留空位情况在此相持续提示 / empty-slot hint kept in this state
        IF (NOT bEnable) OR bReset OR (nEmptySlots = 0 AND (NOT bSpaceWarn)) THEN
            eState := E_DL_CasePackState.eIdle;    // 失能 / 复位 / 无空位提示三条退出条件 / three exits
            IF bReset THEN
                nSeqIndex := DL_CPP_IDX_FIRST;     // 复位沿直接回序号 1 / reset rewinds immediately
            END_IF
        END_IF

    E_DL_CasePackState.eFault:
        bValid := FALSE;                           // 故障闸显式不可用（R72）/ explicit FALSE on the fault gate
        bError := TRUE;                            // 故障级必置 bError（R45 配对）/ fault-class pairs with bError
        nSeqIndex := DL_CPP_IDX_FIRST;             // 故障侧序列回 1，防上层按旧序号取件 / rewind so the upper layer cannot pick on a stale index
        fTargetXMm := DL_CPP_ZERO;                 // 坐标回零安全侧 / coordinates zeroed, safe side
        fTargetYMm := DL_CPP_ZERO;                 // 坐标回零安全侧 / coordinates zeroed, safe side
        fTargetZMm := DL_CPP_ZERO;                 // 坐标回零安全侧 / coordinates zeroed, safe side
        fTargetRotDeg := DL_CPP_ZERO;              // 旋转角回零安全侧 / rotation zeroed, safe side
        bLast := FALSE;                            // 末位标志撤 / last flag withdrawn
        IF eErr = 16#0000_0000 THEN
            eErr := DL_CPP_CODE_FLT_3;             // 入口无码时按非法状态兜底（R45：bError 必须有对应码）/ illegal-state fallback
        END_IF
        IF bEnable AND (nCols >= DL_CPP_DIM_MIN) AND (nCols <= DL_CPP_DIM_MAX)
           AND (nRows >= DL_CPP_DIM_MIN) AND (nRows <= DL_CPP_DIM_MAX)
           AND (nLayers >= DL_CPP_DIM_MIN) AND (nLayers <= DL_CPP_DIM_MAX)
           AND (fPitchXMm > DL_CPP_TOL) AND (fPitchYMm > DL_CPP_TOL) AND (fLayerGapMm > DL_CPP_TOL)
           AND (nBoxCount >= DL_CPP_DIM_MIN) AND (nBoxCount <= nCapacity) THEN
            eState := E_DL_CasePackState.eIdle;    // 全部组态恢复才回待机（退出条件 ≥2）/ recover only when every configuration item is sane
        END_IF

    ELSE
        eState := E_DL_CasePackState.eFault;       // 非法状态兜底 / illegal-state fallback
        eErr := DL_CPP_CODE_FLT_3;                 // 故障级兜底：非法状态 / fault fallback: illegal state
        bError := TRUE;                            // 故障级必置 bError（R45 配对）/ fault-class pairs with bError
        bValid := FALSE;                           // 位姿不可用 / poses unusable
        nSeqIndex := DL_CPP_IDX_FIRST;             // 序列回序号 1 安全侧 / sequence rewound, safe side
        fTargetXMm := DL_CPP_ZERO;                 // 坐标回零安全侧 / coordinates zeroed, safe side
        fTargetYMm := DL_CPP_ZERO;                 // 坐标回零安全侧 / coordinates zeroed, safe side
        fTargetZMm := DL_CPP_ZERO;                 // 坐标回零安全侧 / coordinates zeroed, safe side
        fTargetRotDeg := DL_CPP_ZERO;              // 旋转角回零安全侧 / rotation zeroed, safe side
        bLast := FALSE;                            // 末位标志撤 / last flag withdrawn

END_CASE
END_FUNCTION_BLOCK

(* ---- FB_DL_CasePackerPatternVerify.st ---- *)
(*==============================================================================
 * 组件名称 (Component)  : FB_DL_CasePackerPatternVerify
 * 所属子库 (Sublibrary) : DL_Process
 * 当前版本 (Version)    : 1.0.0
 * 兼容性 (Platform)     : CODESYS 3.5+ / TwinCAT 3 / 汇川 InoProShop / 施耐德 Machine Expert
 *                         仅依赖 Standard.library（R_TRIG），零厂商私有库
 * 功能描述 (Function)   : 装箱排列模式校验防错。装箱到位沿比较传感器位域
 *                         （8 槽）与目标模式字：XOR 全零 → bPatternOk 放行；
 *                         任一位冲突 → bReject 单拍拒启并锁存 bRejectLatch
 *                         给出首错槽位。禁止位掩码 uNoGoMask（重叠占位）置位
 *                         即拒启（重叠即拒启语义）。与 RangeOverlapCheck
 *                         （纯区间函数）分工：本件是模式放行顺控，重叠只是
 *                         拒启判据之一。
 * 来源标签 (Origin)     : ROADMAP §16.4 R11 池（L720），自研 clean-room
 * 边界语义 (Boundary)   : ① 位域冲突 → 首错槽位 1..8 报告，多错只报首个
 *                         （定位修复优先）；
 *                         ② 掩码 SHL 移位量 0..7 < 16 位宽（R48 安全）；
 *                         ③ 拒启锁存至下个到位沿或复位沿（清除路径声明）；
 *                         ④ 无浮点量（纯位域，无 NaN/除零域）。
 * 输出语义 (Fallback)   : 【R191】bEnable = FALSE → 校验输出冻结保持；eFault
 *                         相 → 放行出口强制 FALSE（拒启安全侧）+ bError = TRUE。
 * 码位     (Codes)      : 按 R297 范式零 16# 码位硬编码；错误出口 BOOL+ENUM(eCause)。
 * 红线自检 (Redline)    : 7 项红线已自检：R1 零全局 ✓｜R2 零物理地址 ✓｜R3 纯 IEC ✓
 *                         R4 越界（移位有界）/组态闸 ✓｜R5 双语同行注释 ✓
 *                         R6 CASE 带 ELSE 兜底迁 eFault ✓｜R7 R_TRIG 段 0 无条件刷新 ✓
 * 验收向量 (Acceptance) : V1 uPatternIn=16#00FF、Ref=16#00FF、NoGo=16#0000
 *                         → bPatternOk=TRUE；
 *                         V2 In=16#00FE、Ref=16#00FF → bReject 单拍，首错
 *                         槽位 nErrSlot=8（位 7 对应槽 8）；
 *                         V3 NoGo=16#0001 且 In bit0=1（重叠占位）→ 拒启。
 * 修订历史 (Revision)   : 2026-11-20  v1.0.0  R51 首版（批 2 · 序号 6）
 *==============================================================================*)
TYPE E_DL_CpvState :
(
    eIdle  := 0,                             (* 待使能 / Idle *)
    eArmed := 10,                            (* 武装等待装箱到位沿 / Armed for box edge *)
    eFault := 90                             (* 故障锁存相 / Fault latched phase *)
);
END_TYPE

TYPE E_DL_CpvCause :
(
    eNone     := 0,                          (* 无故障成因 / No cause *)
    ePattern  := 1,                          (* 模式位冲突拒启 / Pattern mismatch reject *)
    eNoGoHit  := 2,                          (* 禁止位（重叠占位）拒启 / No-go overlap reject *)
    ePhaseBad := 3                           (* 非法相位兜底 / Illegal phase fallback *)
);
END_TYPE

FUNCTION_BLOCK FB_DL_CasePackerPatternVerify
VAR_INPUT
    uPatternIn  : WORD := 16#0000;           (* 8 槽传感器位域（1 = 有箱）[-] / Sensor bit field *)
    uPatternRef : WORD := 16#00FF;           (* 目标排列模式字 [-] / Target pattern word *)
    uNoGoMask   : WORD := 16#0000;           (* 禁止位掩码（重叠占位禁放）[-] / No-go mask *)
    bBoxPresent : BOOL := FALSE;             (* 装箱到位电平（上升沿触发校验）[-] / Box present level *)
    bEnable     : BOOL := TRUE;              (* 使能 [-] / Enable *)
    bReset      : BOOL := FALSE;             (* 复位命令，上升沿清全部 [-] / Reset command *)
END_VAR
VAR_OUTPUT
    bPatternOk  : BOOL;                      (* 模式匹配放行（校验拍保持到下个沿）[-] / Pattern pass *)
    bReject     : BOOL;                      (* 拒启单拍位 [-] / Reject pulse *)
    bRejectLatch: BOOL;                      (* 拒启锁存（下个到位沿或复位沿清）[-] / Reject latch *)
    nErrSlot    : INT;                       (* 首错槽位 1..8（无错为 0）[槽] / First error slot *)
    nVerifyCnt  : UDINT;                     (* 累计校验次数 [次] / Verify count *)
    eState      : E_DL_CpvState;             (* 状态出口 / State outlet *)
    eCause      : E_DL_CpvCause;             (* 故障成因出口（R190 独立分码） / Fault cause outlet *)
    bError      : BOOL;                      (* 故障锁存标志 [-] / Fault latch flag *)
END_VAR
VAR
    _eState    : E_DL_CpvState := E_DL_CpvState.eIdle;     (* 内部相位（CASE 唯一写入目标） / Internal phase *)
    _eCause    : E_DL_CpvCause := E_DL_CpvCause.eNone;     (* 故障成因锁存量 / Latched cause *)
    rtBox      : R_TRIG;                     (* 到位沿实例，段 0 无条件调用 / Box edge instance *)
    rtReset    : R_TRIG;                     (* 复位沿实例，段 0 无条件调用 / Reset edge instance *)
    _wDiff     : WORD;                       (* 异或差掩码工作量 [-] / XOR diff work *)
    _bPass     : BOOL;                       (* 放行锁存 [-] / Pass latch *)
    _nSlot     : INT;                        (* 首错槽位锁存 [槽] / First-error slot latch *)
    _i         : INT;                        (* 槽扫描游标（每趟重置，R227）[-] / Slot cursor *)
    _wMask     : WORD;                       (* 槽位掩码工作量 [-] / Slot mask work *)
    _nVerC     : UDINT;                      (* 校验计数锁存 [次] / Verify count latch *)
    _bFault    : BOOL;                       (* 故障锁存位 / Latched fault bit *)
END_VAR
VAR CONSTANT
    DL_CPV_SLOTS : INT := 8;                 (* 槽位总数 [槽] / Slot count *)
END_VAR

(* —— 段 0：沿实例无条件刷新（R228A；纯位域件无浮点组态闸） —— *)
rtBox(CLK := bBoxPresent);                   (* 到位沿每拍必调 / Box edge every scan *)
rtReset(CLK := bReset);                      (* 复位沿每拍必调 / Reset edge every scan *)

(* —— 段 1：单拍量预清零（R107） —— *)
bReject := FALSE;                            (* 拒启脉冲预清，唯一分支置位 / Reject preset *)

(* —— 段 2：复位沿处理（作用域：清故障 + 清锁存 + 清出口 + 清计数 + 迁 eIdle，R283 逐项声明） —— *)
IF rtReset.Q THEN
    _bFault := FALSE;                        (* 清故障锁存 / Clear fault *)
    _eCause := E_DL_CpvCause.eNone;          (* 清成因 / Clear cause *)
    _bPass := FALSE;                         (* 清放行锁存 / Clear pass latch *)
    bRejectLatch := FALSE;                   (* 清拒启锁存 / Clear reject latch *)
    _nSlot := 0;                             (* 清首错槽 / Clear slot *)
    nErrSlot := 0;                           (* 清槽位出口 / Clear slot outlet *)
    bPatternOk := FALSE;                     (* 清放行出口 / Clear pass outlet *)
    _nVerC := 0;                             (* 清校验计数 / Clear count *)
    _eState := E_DL_CpvState.eIdle;          (* 迁待机相 / Back to idle *)
END_IF

(* —— 段 4：CASE 主状态机（ELSE 兜底迁 eFault，红线 6；无组态浮点闸故无段 3） —— *)
CASE _eState OF
    E_DL_CpvState.eIdle:                     (* 待机相 / Idle *)
        IF bEnable AND NOT _bFault THEN
            _eState := E_DL_CpvState.eArmed; (* 进入武装 / Enter armed *)
        END_IF
    E_DL_CpvState.eArmed:                    (* 武装相：到位沿校验 / Armed *)
        IF NOT bEnable THEN
            _eState := E_DL_CpvState.eIdle;  (* 失能回待机 / Back to idle *)
        ELSIF rtBox.Q THEN                   (* 到位沿：执行校验 / Verify on edge *)
            _nVerC := _nVerC + 1;            (* 校验计数（UDINT 回绕工程安全） / Count verify *)
            IF (uPatternIn AND uNoGoMask) <> 16#0000 THEN   (* 禁止位命中：重叠占位拒启（R190 独立分码） / No-go overlap hit *)
                _eCause := E_DL_CpvCause.eNoGoHit;   (* 成因：重叠 / Cause: overlap *)
                _bFault := TRUE;             (* 故障锁存（R45 配对：出口由段 5 强制拒启） / Latch fault *)
                _eState := E_DL_CpvState.eFault;   (* 迁故障相 / To fault *)
                bReject := TRUE;             (* 拒启单拍 / Reject pulse *)
                bRejectLatch := TRUE;        (* 拒启锁存 / Reject latch *)
            ELSE
                _wDiff := uPatternIn XOR uPatternRef;   (* 异或差掩码 / XOR diff *)
                IF _wDiff = 16#0000 THEN
                    _bPass := TRUE;          (* 全零匹配放行 / Pass *)
                    bPatternOk := TRUE;      (* 放行出口 / Pass outlet *)
                    _nSlot := 0;             (* 无错清槽 / Clear slot *)
                    nErrSlot := 0;           (* 槽位出口清 / Slot outlet clear *)
                    bRejectLatch := FALSE;   (* 此前拒启锁存清除（到位沿清除路径，边界③） / Clear reject latch *)
                ELSE
                    _i := 0;                 (* 槽游标重置（R227） / Slot cursor reset *)
                    _wMask := 16#0001;       (* 掩码起点（位 0 = 槽 1） / Mask start *)
                    _nSlot := 0;             (* 首错槽预置 0 / Slot preset *)
                    WHILE (_i <= DL_CPV_SLOTS - 1) AND (_nSlot = 0) DO   (* 逐槽找首错（移位量 0..7 < 16，R48） / First error slot *)
                        IF (_wDiff AND _wMask) <> 16#0000 THEN
                            _nSlot := _i + 1;   (* 槽号 = 位号 + 1 / Slot number *)
                        END_IF
                        _wMask := SHL(_wMask, 1);   (* 掩码左移（常量 1 位） / Shift mask *)
                        _i := _i + 1;        (* 游标递进 / Cursor advance *)
                    END_WHILE
                    _eCause := E_DL_CpvCause.ePattern;   (* 成因：模式冲突 / Cause: pattern *)
                    _bFault := TRUE;         (* 故障锁存（R45 配对） / Latch fault *)
                    _eState := E_DL_CpvState.eFault;   (* 迁故障相 / To fault *)
                    nErrSlot := _nSlot;      (* 首错槽出口 / Slot outlet *)
                    bReject := TRUE;         (* 拒启单拍 / Reject pulse *)
                    bRejectLatch := TRUE;    (* 拒启锁存 / Reject latch *)
                END_IF
            END_IF
        END_IF
    E_DL_CpvState.eFault:                    (* 故障相：放行出口强制 FALSE（安全侧），仅复位沿出 / Fault *)
        bPatternOk := FALSE;                 (* 放行收敛 / Pass converge *)
    ELSE                                     (* 非法相位兜底迁安全态 / Illegal phase fallback *)
        _eState := E_DL_CpvState.eFault;     (* 迁故障相 / To fault *)
        _bFault := TRUE;                     (* 同步锁存 / Latch *)
        _eCause := E_DL_CpvCause.ePhaseBad;  (* 成因：非法相位 / Cause: illegal phase *)
END_CASE

(* —— 段 5：出口映射（bError/eState 同源，R191） —— *)
nVerifyCnt := _nVerC;                        (* 校验计数出口 / Count outlet *)
bError := _bFault;                           (* 故障标志镜像 / Fault flag mirror *)
eState := _eState;                           (* 状态出口 / State outlet *)
eCause := _eCause;                           (* 成因出口 / Cause outlet *)
END_FUNCTION_BLOCK

(* ---- FB_DL_CaseSealerFlapFoldSeq.st ---- *)
(*==============================================================================
 * 组件名称 (Component)  : FB_DL_CaseSealerFlapFoldSeq
 * 所属子库 (Sublibrary) : DL_Process
 * 归属目录 (Directory)  : C:\Library\DL_Process
 * 当前版本 (Version)    : 1.0.0
 * 分类/来源标签         : 功能块（FUNCTION_BLOCK）· 包装机械 · 封箱机折盖顺控
 *                         industry-pool / packaging / case-sealer / sequence
 * 兼容性   (Platform)   : CODESYS 3.5 / TwinCAT 3 / 汇川 InoProShop / 施耐德
 *                         Machine Expert；仅用 Standard.library 的 TON / R_TRIG
 * 溯源声明 (Provenance) : 道莅自研 clean-room——只借公开规范条款与工程惯例，零代码行复制。
 * 功能一句话 (Summary)  : 封箱机折盖六步顺控：进箱确认 → 折后盖 → 折前盖 →
 *                         压盖封箱（胶带/热熔双模式抽象）→ 完成，步序守护超时。
 *
 * 功能描述 (Function)   : 步进状态机：每步以到位传感器为转移条件，每步独立
 *                         守护超时（单步超时即卡箱故障，冻结输出保守停机）；
 *                         封箱步按模式区分：胶带模式只压盖，热熔模式压盖
 *                         加热熔 dwell 计时；完成以信息级 3028 告知并回待机。
 *                         箱未到位禁止起步折页（联锁拒绝），非法状态拦截。
 * 与既有件边界 (Boundary): 进箱/出箱输送线控制归输送件；本件只编排折盖
 *                         与封箱动作，不驱动输送。
 * 码位说明 (Codes)      : 信息 16#0006_3028 一箱封箱完成
 *                         故障 16#0006_3029 步序守护超时，卡箱保守停机
 *                         故障 16#0006_302A 箱未到位禁止起步（联锁拒绝）
 *                         故障 16#0006_302B 封箱模式域外
 *                         段 16#06_0_28~2C 首槽信息级、次槽起故障级。
 * 依赖说明 (Depends)    : 无 DL_ 内部依赖；仅 Standard.library 的 TON / R_TRIG。
 * 红线自检 (Redline)    : 零全局依赖 ｜ 零 VAR_EXTERNAL ｜ 零 %I/%Q（输出引脚）
 *                         TON/R_TRIG 每周期无条件刷新 ｜ ENUM 配 CASE 且 ELSE 兜底
 *                         多段守护用 ARRAY[1..6] OF TON 独立实例（R158）
 *                         全变量双语同行注释 ｜ 故障锁存回放且有可达解除路径
 * 修订历史 (Revision)   : 2026-11-18  v1.0.0  首版入库（R32 · 批 4）
 *============================================================================*)

FUNCTION_BLOCK FB_DL_CaseSealerFlapFoldSeq
VAR_INPUT
    bRun         : BOOL;                // 顺控使能，假则回待机 / Enable, FALSE stands by
    bBoxPresent  : BOOL;                // 箱到位传感器 [开关] / Box present sensor
    bFlapRearFwd : BOOL;                // 后盖折页到位 [开关] / Rear flap folded sensor
    bFlapFrontFwd: BOOL;                // 前盖折页到位 [开关] / Front flap folded sensor
    bPressFwd    : BOOL;                // 压盖缸到位 [开关] / Press cylinder forward sensor
    eSealMode    : (eTape := 0, eHotMelt := 1); // 封箱模式枚举：胶带/热熔 / Seal mode enum
    tStepGuard   : TIME  := T#10S;      // 单步守护超时 [s] / Per-step guard timeout
    tDwellHM     : TIME  := T#2S;       // 热熔 dwell 时长 [s] / Hot-melt dwell duration
END_VAR
VAR_OUTPUT
    oFoldRear: BOOL;                    // 后盖折页缸输出 [引脚] / Rear flap cylinder output
    oFoldFront: BOOL;                   // 前盖折页缸输出 [引脚] / Front flap cylinder output
    oPressCyl: BOOL;                    // 压盖缸输出 [引脚] / Press cylinder output
    oSealAct : BOOL;                    // 封箱动作输出（胶带贴附或热熔加热）[引脚] / Seal action output
    eStep    : (eStStandby := 0, eStFoldRear := 1, eStFoldFront := 2, eStPress := 3, eStDwell := 4, eStDone := 5);   // 步序枚举输出 / Step output enum
    bDone    : BOOL;                    // 一箱完成脉冲 [事件] / One-shot box done pulse
    bError   : BOOL;                    // 故障标志，与故障码配对 / Fault flag paired with codes
    uErrorId : UDINT;                   // 事件码，0 表示无事件 / Event code, zero means none
END_VAR
VAR
    _eStep    : (eStStandby := 0, eStFoldRear := 1, eStFoldFront := 2, eStPress := 3, eStDwell := 4, eStDone := 5);  // 内部步序 / Internal step
    aTonGuard : ARRAY[1..6] OF TON;     // 各步守护定时器（R158 独立实例）/ Per-step guard timers
    tonDwell  : TON;                    // 热熔 dwell 定时器 [s] / Hot-melt dwell timer
    rTrigBox  : R_TRIG;                 // 箱到位上升沿 / Box present rising edge
    bGuardAct : BOOL;                   // 守护超时锁存 / Guard timeout latched
    uCodeLatch: UDINT;                  // 故障锁存码 [码] / Latched fault code
    uInfoCode : UDINT;                  // 信息级单拍码 [码] / One-shot info code
END_VAR
VAR CONSTANT
    DL_CSF_NSTEPS : INT := 6;           // 步数 [步]，与数组声明一致 / Step count, matches the array
END_VAR

(* 段 1｜定时器与边沿无条件刷新（红线 7）：六步守护独立实例 + dwell + 箱沿
 *      Timers refreshed unconditionally: six per-step guards, dwell, box edge *)
bGuardAct := FALSE;                     // 守护标志本拍重估 / Re-evaluate this scan
rTrigBox(CLK := bBoxPresent);           // 箱到位沿检测 / Box edge detection
tonDwell(IN := (_eStep = eStDwell), PT := tDwellHM);    // dwell 计时 / Dwell timing

(* 段 2｜六步守护矩阵：六实例每拍无条件刷新（R158）/ Guard matrix, six instances refreshed every scan *)
aTonGuard[1](IN := (_eStep = eStStandby)  AND bRun, PT := tStepGuard);
aTonGuard[2](IN := (_eStep = eStFoldRear) AND bRun, PT := tStepGuard);
aTonGuard[3](IN := (_eStep = eStFoldFront) AND bRun, PT := tStepGuard);
aTonGuard[4](IN := (_eStep = eStPress)    AND bRun, PT := tStepGuard);
aTonGuard[5](IN := (_eStep = eStDwell)    AND bRun, PT := tStepGuard);
aTonGuard[6](IN := (_eStep = eStDone)     AND bRun, PT := tStepGuard);
bGuardAct := aTonGuard[2].Q OR aTonGuard[3].Q OR aTonGuard[4].Q OR aTonGuard[5].Q;  // 任一活动步超时 / Any active step timed out
IF bGuardAct THEN
    uCodeLatch := 16#0006_3029;         // 故障级：步序守护超时 / Fault: step guard timeout
END_IF

(* 段 3｜步进状态机主分派（ENUM 配 CASE，ELSE 兜底）/ Step dispatch with ELSE interception *)
CASE _eStep OF

    eStStandby:
        (* 本拍行为：全输出撤；使能与箱到位俱备拍 N+1 起步 / All off; start on box present *)
        oFoldRear := FALSE;             // 撤后盖缸 / Retract the rear cylinder
        oFoldFront := FALSE;            // 撤前盖缸 / Retract the front cylinder
        oPressCyl := FALSE;             // 撤压盖缸 / Retract the press
        oSealAct := FALSE;              // 撤封箱动作 / Withdraw the seal action
        bDone := FALSE;                 // 完成脉冲清 / Clear the done pulse
        IF bRun AND rTrigBox.Q THEN
            _eStep := eStFoldRear;      // 拍 N+1 起步折后盖 / To fold rear next scan
        END_IF

    eStFoldRear:
        (* 本拍行为：驱动后盖缸；到位转折前盖 / Drive the rear cylinder; transfer on sensor *)
        oFoldRear := TRUE;              // 驱动后盖 / Drive the rear
        oFoldFront := FALSE;
        oPressCyl := FALSE;
        oSealAct := FALSE;
        IF NOT bRun THEN
            _eStep := eStStandby;       // 撤使能回待机 / Disable to standby
        ELSIF bFlapRearFwd THEN
            _eStep := eStFoldFront;     // 拍 N+1 转折前盖 / To fold front next scan
        END_IF

    eStFoldFront:
        (* 本拍行为：驱动前盖缸；到位转压盖 / Drive the front cylinder *)
        oFoldRear := FALSE;
        oFoldFront := TRUE;             // 驱动前盖 / Drive the front
        oPressCyl := FALSE;
        oSealAct := FALSE;
        IF NOT bRun THEN
            _eStep := eStStandby;       // 撤使能回待机 / Disable to standby
        ELSIF bFlapFrontFwd THEN
            _eStep := eStPress;         // 拍 N+1 转压盖 / To press next scan
        END_IF

    eStPress:
        (* 本拍行为：压盖缸进；到位后按模式转封箱动作或 dwell / Press; transfer by mode *)
        oFoldRear := FALSE;
        oFoldFront := FALSE;
        oPressCyl := TRUE;              // 驱动压盖 / Drive the press
        oSealAct := FALSE;
        IF NOT bRun THEN
            _eStep := eStStandby;       // 撤使能回待机 / Disable to standby
        ELSIF bPressFwd THEN
            CASE eSealMode OF           // 模式内嵌 CASE（枚举配 ELSE）/ Nested mode CASE with ELSE
                eTape:    _eStep := eStDone;    // 胶带模式：压盖即完成 / Tape: press is enough
                eHotMelt: _eStep := eStDwell;   // 热熔模式：转 dwell / Hot melt: dwell
            ELSE
                uCodeLatch := 16#0006_302B;     // 故障级：模式域外 / Fault: mode out of range
                _eStep := eStStandby;
            END_CASE
        END_IF

    eStDwell:
        (* 本拍行为：压盖保持 + 封箱动作输出，dwell 满完成 / Hold and seal, done on dwell *)
        oFoldRear := FALSE;
        oFoldFront := FALSE;
        oPressCyl := TRUE;              // 保持压盖 / Hold the press
        oSealAct := TRUE;               // 热熔加热输出 / Hot melt output
        IF NOT bRun THEN
            _eStep := eStStandby;       // 撤使能回待机 / Disable to standby
        ELSIF tonDwell.Q THEN
            _eStep := eStDone;          // dwell 满，拍 N+1 完成 / Done next scan
        END_IF

    eStDone:
        (* 本拍行为：全输出撤 + 完成脉冲单拍，箱离位回待机 / All off, one-shot pulse, wait for box leave *)
        oFoldRear := FALSE;
        oFoldFront := FALSE;
        oPressCyl := FALSE;
        oSealAct := FALSE;
        bDone := TRUE;                  // 完成脉冲（单拍）/ One-shot done pulse
        uInfoCode := 16#0006_3028;      // 信息级：一箱完成 / Info: box done
        IF NOT bBoxPresent THEN
            _eStep := eStStandby;       // 箱离位回待机 / Box left, to standby
        END_IF
        IF NOT bRun THEN
            _eStep := eStStandby;       // 撤使能回待机 / Disable to standby
        END_IF

ELSE
    oFoldRear := FALSE;                 // 非法步全撤（保守停机）/ Illegal step, all off
    oFoldFront := FALSE;
    oPressCyl := FALSE;
    oSealAct := FALSE;
    _eStep := eStStandby;               // 拦截回待机 / Intercept to standby
    uCodeLatch := 16#0006_3029;         // 故障：步序越界 / Fault: step out of range
END_CASE

(* 段 4｜出口装配 / Exit assembly *)
eStep := _eStep;                        // 步序枚举输出 / Step output
IF NOT bRun THEN
    uCodeLatch := 16#0000_0000;         // 撤使能清故障（可达解除）/ Run drop clears faults
END_IF
bError := (uCodeLatch <> 16#0000_0000); // 故障锁存回放 / Latched fault replay
IF uCodeLatch <> 16#0000_0000 THEN
    uErrorId := uCodeLatch;             // 故障码优先 / Fault first
    uInfoCode := 16#0000_0000;
ELSE
    uErrorId := uInfoCode;              // 信息码单拍 / Info one shot
    uInfoCode := 16#0000_0000;
END_IF
END_FUNCTION_BLOCK

(* ---- FB_DL_CaseShiftTally.st ---- *)
(*
  Name        : FB_DL_CaseShiftTally
  Category    : DL_Process
  Version     : 1.0.0
  Purpose     : 班次箱数台账与计划差异告警：班次激活期逐箱计数，班末与计划量比对，偏差百分比超容差即告警并保持至下班次启动；/ Shift case tally with plan-deviation alarm: counts cases while the shift is active, compares against plan at shift end, alarms when deviation exceeds tolerance and holds until the next shift starts
  溯源        : 借 ROADMAP P2（BidirectionalCounter/OeeCalculator 口径复用），clean-room 实现
  Boundary    : ① 组态闸：计划量 < 1 / 容差 < 0 → 锁存故障（计划量 0 使偏差比无定义）；
                ② 除零前置：偏差比除子为计划量，组态闸保证 >= 1；
                ③ 计数仅在 eCount 相（班次激活）沿触发累加，班末（bShiftEnd 沿）一次性结算；
                ④ 台账语义：eDone 相保持 nActual/fDevPct/bDevAlarm 电平（锁存副本），不随实时量回落（族② 口径）；
                ⑤ 下班次 bShiftStart 沿清台账开新班（唯一清零路径，另有复位沿全清）；
                ⑥ 本件只做台账与告警，不执行停机（属主边界）。
*)
TYPE E_DL_CstState :
(
    eIdle  := 0,                             (* 待班次启动 / Waiting shift start *)
    eCount := 10,                            (* 班次计数中 / Counting *)
    eDone  := 20,                            (* 班末结算完成（保持台账） / Settled, tally held *)
    eFault := 90                             (* 故障锁存相 / Fault latched *)
);
END_TYPE

TYPE E_DL_CstCause :
(
    eNone       := 0,                        (* 无故障成因 / No cause *)
    eCfgIllegal := 1,                        (* 组态非法：计划量/容差越域 / Illegal config *)
    ePhaseBad   := 2                         (* 非法相位兜底 / Illegal phase fallback *)
);
END_TYPE

FUNCTION_BLOCK FB_DL_CaseShiftTally
VAR_INPUT
    bCasePass   : BOOL := FALSE;             (* 单箱过站脉冲（上升沿计一箱）[-] / One case passed pulse *)
    nPlanQty    : UDINT := 100;              (* 班次计划箱数，域 >= 1 [箱] / Planned case quantity, >= 1 *)
    fTolPct     : REAL := 10.0;              (* 偏差告警容差，域 >= 0 [%] / Deviation tolerance, >= 0 *)
    bShiftActive: BOOL := FALSE;             (* 班次激活电平（计数的门控条件）[-] / Shift active level *)
    bShiftStart : BOOL := FALSE;             (* 班次启动脉冲（清台账开新班）[-] / Shift start pulse *)
    bShiftEnd   : BOOL := FALSE;             (* 班末结算脉冲（一次性比对）[-] / Shift end pulse *)
    bEnable     : BOOL := TRUE;              (* 台账使能 [-] / Enable *)
    bReset      : BOOL := FALSE;             (* 复位命令，上升沿清台账与故障 [-] / Reset command *)
END_VAR
VAR_OUTPUT
    nActual     : UDINT;                     (* 本班实际箱数（eDone 相保持）[箱] / Actual case count, held in done phase *)
    fDevPct     : REAL;                      (* 计划偏差百分比（eDone 相保持）[%] / Plan deviation percentage, held *)
    bDevAlarm   : BOOL;                      (* 偏差超容差告警（eDone 相保持，复位/新班清）[-] / Deviation alarm, held *)
    bSettled    : BOOL;                      (* 班末结算完成电平（eDone 相为 TRUE）[-] / Settled level *)
    eState      : E_DL_CstState;             (* 状态出口 / State outlet *)
    eCause      : E_DL_CstCause;             (* 故障成因出口（R190 归因唯一） / Fault cause outlet *)
    bError      : BOOL;                      (* 故障锁存标志 [-] / Fault latch flag *)
END_VAR
VAR
    _eState  : E_DL_CstState := E_DL_CstState.eIdle;     (* 内部相位（CASE 唯一写入目标） / Internal phase *)
    _eCause  : E_DL_CstCause := E_DL_CstCause.eNone;     (* 故障成因锁存量 / Latched cause *)
    rtCase   : R_TRIG;                       (* 过箱脉冲沿实例，段 0 无条件调用 / Case pulse edge *)
    rtStart  : R_TRIG;                       (* 班次启动沿实例，段 0 无条件调用 / Shift start edge *)
    rtEnd    : R_TRIG;                       (* 班末脉冲沿实例，段 0 无条件调用 / Shift end edge *)
    rtReset  : R_TRIG;                       (* 复位沿实例，段 0 无条件调用 / Reset edge instance *)
    _bFault  : BOOL;                         (* 故障锁存位 / Latched fault bit *)
    _bCfgBad : BOOL;                         (* 组态非法当拍量 / Illegal config this scan *)
    _nCnt    : UDINT;                        (* 本班计数内部量（出口锁存副本源）[箱] / Internal tally, source of held outlet *)
    _fDevI   : REAL;                         (* 偏差比中间量 [%] / Deviation intermediate *)
    _bAlarmI : BOOL;                         (* 告警内部量（锁存副本源）[-] / Alarm internal, source of held outlet *)
    _fSign   : REAL;                         (* 偏差方向符号中间量（+超产/-欠产）[-] / Deviation sign intermediate *)
END_VAR
VAR CONSTANT
    DL_CST_EPS    : REAL  := 1.0E-6;         (* 判零容差 [-] / Epsilon *)
    DL_CST_CNTMAX : UDINT := 4294967295;     (* 计数饱和上限（R28）[-] / Count saturation cap *)
    DL_CST_HUND   : REAL  := 100.0;          (* 百分数换算常量（乘性常量）[-] / Percent scale constant *)
END_VAR

(* —— 段 0：当拍判据派生 + 实例无条件刷新（R228A；四 R_TRIG 全在段 0，无 IF 包裹） —— *)
_bCfgBad := (nPlanQty < 1) OR (fTolPct < 0.0);                                 (* 计划量下限闸 + 容差非负闸 / Plan and tolerance gates *)
rtCase(CLK := bCasePass);                                                      (* 过箱沿每拍必调 / Case edge every scan *)
rtStart(CLK := bShiftStart);                                                   (* 班启动沿每拍必调 / Start edge every scan *)
rtEnd(CLK := bShiftEnd);                                                       (* 班末沿每拍必调 / End edge every scan *)
rtReset(CLK := bReset);                                                        (* 复位沿每拍必调 / Reset edge every scan *)

(* —— 段 1：单拍量预清零（R107；nActual/fDevPct/bDevAlarm 为锁存出口，不在此预清，族② 口径） —— *)
_bAlarmI := FALSE;                                                             (* 告警内部量预清（结算拍重算） / Alarm internal preset *)
_fDevI := 0.0;                                                                 (* 偏差中间量预清 / Deviation preset *)
_fSign := 1.0;                                                                 (* 方向符号预置（默认超产方向） / Sign preset *)

(* —— 段 2：复位沿处理（作用域：清故障 + 清台账 + 迁 eIdle，R283 逐项声明） —— *)
IF rtReset.Q THEN
    _bFault := FALSE;                                                          (* 清故障锁存 / Clear fault *)
    _eCause := E_DL_CstCause.eNone;                                            (* 清成因 / Clear cause *)
    _nCnt := 0;                                                                (* 清计数内部量 / Clear tally internal *)
    nActual := 0;                                                              (* 清实际数出口 / Clear actual outlet *)
    fDevPct := 0.0;                                                            (* 清偏差出口 / Clear deviation outlet *)
    bDevAlarm := FALSE;                                                        (* 清告警出口 / Clear alarm outlet *)
    bSettled := FALSE;                                                         (* 清结算电平出口 / Clear settled outlet *)
    _eState := E_DL_CstState.eIdle;                                            (* 迁待班相 / Back to idle *)
END_IF

(* —— 段 3：组态故障锁存（锁存至复位沿，R189） —— *)
IF _bCfgBad AND NOT _bFault THEN
    _bFault := TRUE;                                                           (* 锁存故障位 / Latch fault *)
    _eCause := E_DL_CstCause.eCfgIllegal;                                      (* 成因：组态非法 / Cause: illegal config *)
    _eState := E_DL_CstState.eFault;                                           (* 同步迁故障相 / Migrate to fault *)
END_IF

(* —— 段 4：CASE 主状态机（ELSE 兜底迁 eFault，红线 6） —— *)
CASE _eState OF
    E_DL_CstState.eIdle:                                                       (* 待班次启动：台账空 / Idle *)
        _nCnt := 0;                                                            (* 待班清计数（防隐性回夹） / Clear tally *)
        nActual := 0;                                                          (* 待班清实际数出口 / Clear actual outlet *)
        fDevPct := 0.0;                                                        (* 待班清偏差出口 / Clear deviation outlet *)
        bDevAlarm := FALSE;                                                    (* 待班清告警出口 / Clear alarm outlet *)
        bSettled := FALSE;                                                     (* 待班清结算电平 / Clear settled outlet *)
        IF bEnable AND NOT _bFault THEN
            IF rtStart.Q THEN                                                  (* 班次启动沿：开新班（唯一清零路径之一） / Shift start edge: open new shift *)
                _nCnt := 0;                                                    (* 新班计数从零起 / New tally from zero *)
                _eState := E_DL_CstState.eCount;                               (* 进计数相 / To counting *)
            END_IF
        END_IF
    E_DL_CstState.eCount:                                                       (* 计数相：班次激活期逐箱累加 / Counting *)
        IF NOT bEnable THEN
            _eState := E_DL_CstState.eIdle;                                    (* 失能回待班（台账清） / Back to idle *)
        ELSE
            IF rtStart.Q THEN                                                  (* 计数中再收启动沿：视为重开班，清零重计 / Restart shift on new start edge *)
                _nCnt := 0;                                                    (* 重开班清零 / Restart from zero *)
            END_IF
            IF rtCase.Q AND bShiftActive THEN                                  (* 班次激活 + 过箱沿：计一箱 / Count on case edge while active *)
                IF _nCnt < DL_CST_CNTMAX THEN
                    _nCnt := _nCnt + 1;                                        (* 计数净额 +1（饱和防回绕，R28） / Net +1, saturated *)
                END_IF
            END_IF
            IF rtEnd.Q THEN                                                    (* 班末沿：一次性结算比对 / Shift end edge: settle once *)
                nActual := _nCnt;                                              (* 实际数出口（锁存副本，eDone 相保持） / Actual outlet, held *)
                _fSign := UDINT_TO_REAL(_nCnt) - UDINT_TO_REAL(nPlanQty);      (* 偏差绝对量（有符号方向）[箱] / Signed deviation *)
                fDevPct := _fSign / UDINT_TO_REAL(nPlanQty) * DL_CST_HUND;     (* 偏差比：除子计划量 >= 1 由组态闸保证 [%] / Deviation ratio, divisor gated *)
                IF ABS(fDevPct) > fTolPct THEN
                    _bAlarmI := TRUE;                                          (* 超容差：告警内部量置位 / Over tolerance *)
                END_IF
                bDevAlarm := _bAlarmI;                                         (* 告警出口（锁存副本，保持至新班/复位） / Alarm outlet, held *)
                bSettled := TRUE;                                              (* 结算完成电平置位 / Settled level *)
                _eState := E_DL_CstState.eDone;                                (* 迁完成相（保持台账） / To done *)
            END_IF
        END_IF
    E_DL_CstState.eDone:                                                        (* 完成相：保持台账至下班次启动（族② 保持语义） / Done: hold tally *)
        IF NOT bEnable THEN
            _eState := E_DL_CstState.eIdle;                                    (* 失能回待班（出口随 eIdle 清） / Back to idle *)
        ELSIF rtStart.Q THEN                                                   (* 新班启动沿：清台账重开（唯一保持出口路径） / New shift: clear and restart *)
            _nCnt := 0;                                                        (* 新班计数从零起 / New tally from zero *)
            nActual := 0;                                                      (* 清实际数出口 / Clear actual outlet *)
            fDevPct := 0.0;                                                    (* 清偏差出口 / Clear deviation outlet *)
            bDevAlarm := FALSE;                                                (* 清告警出口 / Clear alarm outlet *)
            bSettled := FALSE;                                                 (* 清结算电平 / Clear settled outlet *)
            _eState := E_DL_CstState.eCount;                                   (* 进新班计数相 / To counting *)
        END_IF
    E_DL_CstState.eFault:                                                       (* 故障相：冻结保持末值，仅复位沿出 / Fault *)
        ;                                                                      (* 锁存回放（R28） / Replay from latch *)
    ELSE                                                                       (* 非法相位兜底迁安全态 / Illegal phase fallback *)
        _eState := E_DL_CstState.eFault;                                       (* 迁故障相 / To fault *)
        _bFault := TRUE;                                                       (* 同步锁存 / Latch *)
        _eCause := E_DL_CstCause.ePhaseBad;                                    (* 成因：非法相位 / Cause: illegal phase *)
END_CASE

(* —— 段 5：出口映射（bError/eState 同源，R191） —— *)
bError := _bFault;                                                             (* 故障标志镜像 / Fault flag mirror *)
eState := _eState;                                                             (* 状态出口 / State outlet *)
eCause := _eCause;                                                             (* 成因出口 / Cause outlet *)
END_FUNCTION_BLOCK

(* ---- FB_DL_CassetteMapVerify.st ---- *)
(*
  FB_DL_CassetteMapVerify  —  花篮片位映射比对校验（Mapping 序列解析 + 错片定位） / Cassette slot-map verify with first-error slot location
  分类 Category : DL_Process
  版本 Version  : 1.0.1
  兼容性 Platform: CODESYS 3.5 / TwinCAT 3 / 汇川 InoProShop / Machine Expert（仅 Standard.library）
  来源 Source   : roadmap-semi-p2 — 半导体花篮 Mapping 缺口件（与 WaferCassetteSlot 槽位监视分工：那件管槽位实时态，本件管映射比对校验）
  溯源 Origin   : clean-room 实现，未复制任何源码行
  功能 Function : 1) 8 槽映射比对：bVerifyCmd 沿承载，wErrMap := wExpMap XOR
                  wActMap（异或位图逐槽比对），wErrMap = 16#0000 → 校验通过
                  （信息级 04B9）；非零 → 0391 映射失配锁存 + 首错槽位定位
                  （nFirstErrSlot 取最低错位槽号，信息级 04BB）；
                  2) 组态闸：wExpMap = 16#0000（空花篮无校验意义）→ 0392 锁存；
                  3) 相位机：eIdle → eDone（比对完成稳态）→ eFault；错片定位
                  只在失配沿承载一次，锁存期不重扫（禁按当下输入重推断）；
                  4) 信息级三码：校验通过 / 失配检出 / 首错定位（沿置位，复位沿
                  清除——v1.0.1 按信息码复位沿清除范式收敛，原单拍沿改锁存）；
                  5) 解除式全当拍量（R240 落地），逐 BOOL 标注见段 4。
  边界 Boundary : ① 槽位掩码 SHL(WORD#1, 0..7)，移位量域 < 16 结构性安全（R48）；
                  ② wActMap 信任来源为槽位传感器组态（头注释声明信任边界）；
                  ③ 失配锁存码由锁存回放，不随后续 wActMap 漂移（R152 回放纪律）；
                  ④ 零全局耦合：无全局变量表依赖、无外部变量声明、无物理 IO 地址。
  依赖 Depends  : Standard.library（R_TRIG）
  码表 Error codes（Process 段 0005，窗口 0391~0393 / 04B9~04BB）:
    16#0005_0391 故障级：映射失配锁存（首错槽号入 nFirstErrSlot），锁存至 bReset
    16#0005_0392 故障级：组态非法（期望图 16#0000 空花篮无效），锁存至 bReset
    16#0005_0393 故障级：相位落 ELSE 兜底，锁存至 bReset
    16#0005_04B9 信息级：校验通过（沿置位，复位沿清除）
    16#0005_04BA 信息级：失配检出（沿置位，复位沿清除）
    16#0005_04BB 信息级：首错槽位定位（nFirstErrSlot 写定拍置位，复位沿清除）
  修订历史 Revision :
    2026-11-19  v1.0.0  R42 首版（批次 3 · 序号 2）
    2026-11-19  v1.0.1  R44 P0 返修（R43 挂账 3 条）：①信息码复位沿清除范式——
                        原实现 _uInfo 每拍重算致 04B9/04BA/04BB 单拍即逝且 HMI 不可
                        采样，借用 FB_DL_DeviceParamVerify v1.0.1 修法改为锁存至
                        bReset 上升沿清除（段 1 预清零撤销、两处解除沿补清）；
                        ②锁存解除式可达自证复核——rtReset.Q 输入引脚当拍量恒可达，
                        维持原解除式不动；③R228A 补查——rtVerify/rtReset 段 0 无条件
                        刷新在位、本件无 TON 实例，补查通过零改动；无关逻辑零改动。
*)

TYPE E_DL_CmvState :
(
    eIdle   := 0,    // 空闲：等校验指令 / Idle, waiting verify command
    eDone   := 10,   // 完成：比对稳态（通过） / Done, verified steady
    eFault  := 90    // 故障：失配或组态锁定 / Fault, latched
);
END_TYPE

FUNCTION_BLOCK FB_DL_CassetteMapVerify
VAR_INPUT
    wExpMap      : WORD := 16#00FF;   // 期望映射位图，位 n = 槽 n 有片 [-] / Expected slot map bitmap
    wActMap      : WORD := 16#00FF;   // 实际映射位图（槽位传感器组态）[-] / Actual slot map bitmap
    bVerifyCmd   : BOOL := FALSE;     // 校验指令，上升沿承载比对 [-] / Verify command edge
    bReset       : BOOL := FALSE;     // 复位，上升沿清故障锁存 / Reset edge clears fault latch
END_VAR
VAR_OUTPUT
    eState       : E_DL_CmvState;     // 状态出口，段尾单点映射 / State outlet
    wErrMap      : WORD;              // 失配位图镜像（异或结果，锁存快照）/ Mismatch bitmap snapshot
    nFirstErrSlot: DINT;              // 首错槽号 [0..7]，-1 = 无首错 / First error slot index
    bMatch       : BOOL;              // 比对通过标志（eDone 相电平）[-] / Match flag
    bError       : BOOL;              // 故障锁存标志 / Fault latch flag
    nErrId       : UDINT;             // 事件码，0 = 无事件 / Event code
END_VAR
VAR
    rtVerify     : R_TRIG;            // 校验指令沿实例，无条件刷新 / Verify edge instance
    rtReset      : R_TRIG;            // 复位沿实例，无条件刷新 / Reset edge instance
    _eState      : E_DL_CmvState := E_DL_CmvState.eIdle;  // 内部相位（CASE 唯一写入目标）/ Internal phase
    _nIdx        : DINT;              // 阵列循环索引 [-] / Array loop index
    _bFirstFound : BOOL;              // 首错槽已定位标志（锁存量）/ First-error located flag
    _bFault      : BOOL;              // 故障锁存位（锁存量）/ Latched fault bit
    _uFault      : UDINT;             // 故障码锁存（锁存量）/ Latched fault code
    _uInfo       : UDINT;             // 信息码锁存（沿置位，复位沿清除） / Latched info code
END_VAR

(* —— 段 0：沿实例无条件周期刷新（禁置于 IF/CASE 内） —— *)
rtVerify(CLK := bVerifyCmd);         // 校验沿（每拍必调）
rtReset(CLK := bReset);              // 复位沿（每拍必调）

(* —— 段 1：单拍量预清零（锁存量 _bFault/_uFault/_bFirstFound/_uInfo/wErrMap 不入清单，
     禁同拍抹除；信息码 v1.0.1 起为锁存量，仅复位沿清除） —— *)
bMatch := FALSE;                    // 通过标志缺省 FALSE
nErrId := 16#0000_0000;             // 事件码缺省无事件

(* —— 段 2：复位沿 + 组态域闸（判据当拍量） —— *)
IF rtReset.Q THEN                   // rtReset.Q = 当拍量
    _bFault := FALSE;               // 清故障锁存位
    _uFault := 16#0000_0000;        // 清故障锁存码
    _uInfo := 16#0000_0000;         // 清信息码锁存（v1.0.1：信息码复位沿清除范式）
    _bFirstFound := FALSE;          // 首错定位标志清零
    nFirstErrSlot := -1;            // 首错槽号恢复哨兵
    wErrMap := 16#0000;             // 失配位图清零
END_IF
IF wExpMap = 16#0000 THEN           // 期望图域闸（空花篮无效，WORD 判等合规）
    _uFault := 16#0005_0392;        // 故障级：组态非法
    _bFault := TRUE;                // 故障标志与码位配对（R45）
END_IF

(* —— 段 3：校验沿承载比对（判据当拍量沿；失配沿单次定位，锁存期不重扫） —— *)
IF rtVerify.Q AND (NOT _bFault) THEN
    wErrMap := wExpMap XOR wActMap; // 异或位图比对（16 位掩码域结构性安全）
    IF wErrMap = 16#0000 THEN
        _uInfo := 16#0005_04B9;     // 信息级：校验通过沿
        _eState := E_DL_CmvState.eDone;     // 进完成稳态相
    ELSE
        _uInfo := 16#0005_04BA;     // 信息级：失配检出沿
        FOR _nIdx := 0 TO 7 DO      // 首错槽定位（自低向高首个错位）
            IF (NOT _bFirstFound) AND ((wErrMap AND SHL(WORD#1, UINT(_nIdx))) <> WORD#0) THEN
                nFirstErrSlot := _nIdx;             // 首错槽号写定（锁存量，仅此处写）
                _bFirstFound := TRUE;               // 定位标志
                _uInfo := 16#0005_04BB;             // 信息级：首错定位沿（覆盖失配沿，后到优先声明）
            END_IF
        END_FOR
        _uFault := 16#0005_0391;    // 故障级：映射失配锁存
        _bFault := TRUE;
        _eState := E_DL_CmvState.eFault;    // 进故障相
    END_IF
END_IF

(* —— 段 4：故障解除式（R240 落地，逐 BOOL 标注）：
     rtReset.Q = 当拍量；NOT bVerifyCmd = 当拍量；wExpMap ≠ 0 为保持量（组态），
     组态修正后配合复位沿当拍量解除，可达。 —— *)
IF rtReset.Q AND (NOT bVerifyCmd) THEN
    _bFault := FALSE;               // 清故障锁存位（锁存量，仅此当拍量解除沿可清）
    _uFault := 16#0000_0000;        // 清故障锁存码（锁存量，仅本当拍量解除沿可清）
    _uInfo := 16#0000_0000;         // 清信息码锁存（v1.0.1：信息码复位沿清除范式）
    _bFirstFound := FALSE;          // 首错定位标志清零（锁存量）
    nFirstErrSlot := -1;            // 首错槽号恢复哨兵
    IF _eState = E_DL_CmvState.eFault THEN
        _eState := E_DL_CmvState.eIdle;     // 故障相迁出：回空闲
    END_IF
END_IF

(* —— 段 5：相位机（CASE 全覆盖 + ELSE 兜底） —— *)
CASE _eState OF

E_DL_CmvState.eIdle:
    ;                               // 空闲：等校验沿（段 3 承载迁出）

E_DL_CmvState.eDone:
    bMatch := TRUE;                 // 通过标志（相电平）
    IF NOT bVerifyCmd THEN          // 校验指令撤销：回空闲（比对结果随相清除）
        _eState := E_DL_CmvState.eIdle;
    END_IF

E_DL_CmvState.eFault:
    ;                               // 故障相：失配锁存回放，等解除沿（段 4 承载迁出）

ELSE
    _uFault := 16#0005_0393;        // 故障级：非法相位兜底
    _bFault := TRUE;
    _eState := E_DL_CmvState.eFault;    // 强制回故障相

END_CASE

(* —— 段 6：出口单点映射（名实同源；锁存码回放，禁同拍抹除） —— *)
IF _bFault THEN
    nErrId := _uFault;              // 故障锁存码回放
    bMatch := FALSE;                // 故障相通过出口强制 FALSE（安全侧）
ELSE
    nErrId := _uInfo;               // 信息码
END_IF
bError := _bFault;                  // 故障标志与锁存位同源
eState := _eState;                  // 状态出口单点映射

END_FUNCTION_BLOCK
